// TIA Portal V20 export
// export: Created 2026-10-20T12:50:57.8913211Z, ExportSetting WithDefaults, DisplayName Totally Integrated Automation Portal, DisplayVersion V20 Update 6, DisplayName TIA Portal Openness, DisplayVersion V20 Update 6, DisplayName TIA Portal Version Control Interface, DisplayVersion V20 Update 6, DisplayName SINAMICS Startdrive Advanced, DisplayVersion V20 SP1, DisplayName SINAMICS Startdrive G130, G150, S120, S150, SINAMICS MV, G220, S200, S210, DisplayVersion V20 SP1, DisplayName SINAMICS Startdrive G110M, G120, G120C, G120D, G120P, G115D, DisplayVersion V20 SP1, DisplayName STEP 7 Professional, DisplayVersion V20 Update 6, DisplayName STEP 7 Safety, DisplayVersion V20 Update 2, DisplayName WinCC Basic/Comfort/Advanced, DisplayVersion V20 Update 6, DisplayName WinCC Unified, DisplayVersion V20 Update 6
FUNCTION_BLOCK "Main_Panel"   // FB16, F_LAD
{ S7_Optimized_Access := 'TRUE' }
VERSION : 0.1
// stored: AutoNumber true, IsIECCheckEnabled false, UDAEnableTagReadback false
   VAR_INPUT
      Estop_Cabinet_Ch1 : Bool;
      Reset_Cabinet : Bool;
      Bypass : "F_Bypass_MainPanel";
   END_VAR
   VAR_OUTPUT
      Safety_OK : Bool;
      Main_Panel_OK : Bool;
      Bypass_Warning : Bool;
      ACK { ExternalAccessible := 'False'; ExternalVisible := 'False'; ExternalWritable := 'False'} : Bool;
   END_VAR
   VAR
      Estop_Cabinet_DB : ESTOP1;
   END_VAR
BEGIN

REGION Network 1: RESET CABINET
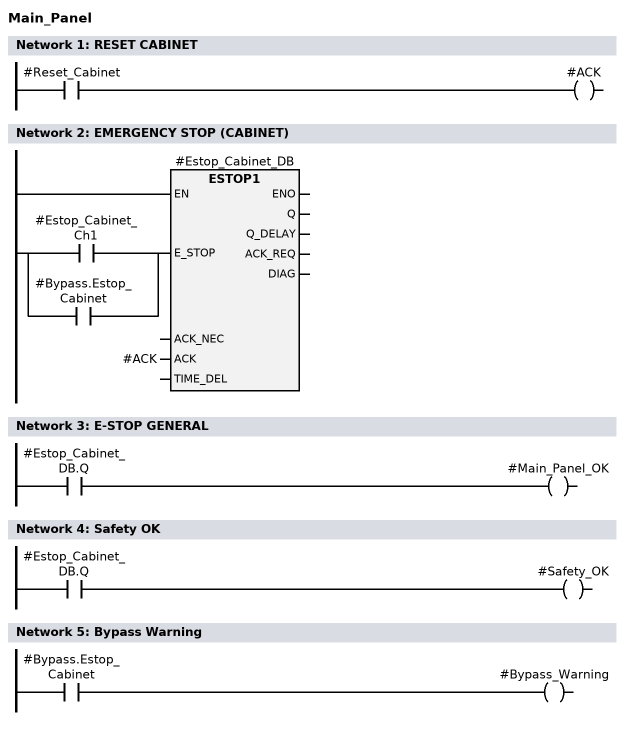
   RUNG wire#powerrail
      Contact( #Reset_Cabinet )
      Coil( #ACK )
   END_RUNG
   // the same network as SCL:
   #ACK := #Reset_Cabinet;
END_REGION

REGION Network 2: EMERGENCY STOP (CABINET)
   RUNG wire#powerrail
      #Estop_Cabinet_DB.ESTOP1(E_STOP := wire#w1, ACK_NEC :=, ACK := #ACK, TIME_DEL :=, Q =>, Q_DELAY =>, ACK_REQ =>, DIAG =>)
   END_RUNG
   RUNG wire#powerrail
      Contact( #Estop_Cabinet_Ch1 )
   END_RUNG wire#w1
   RUNG wire#powerrail
      Contact( #Bypass.Estop_Cabinet )
   END_RUNG wire#w1
   // the same network as SCL:
   #Estop_Cabinet_DB(E_STOP := #Estop_Cabinet_Ch1 OR #Bypass.Estop_Cabinet, ACK := #ACK);   // ESTOP1
END_REGION

REGION Network 3: E-STOP GENERAL
   RUNG wire#powerrail
      Contact( #Estop_Cabinet_DB.Q )
      Coil( #Main_Panel_OK )
   END_RUNG
   // the same network as SCL:
   #Main_Panel_OK := #Estop_Cabinet_DB.Q;
END_REGION

REGION Network 4: Safety OK
   RUNG wire#powerrail
      Contact( #Estop_Cabinet_DB.Q )
      Coil( #Safety_OK )
   END_RUNG
   // the same network as SCL:
   #Safety_OK := #Estop_Cabinet_DB.Q;
END_REGION

REGION Network 5: Bypass Warning
   RUNG wire#powerrail
      Contact( #Bypass.Estop_Cabinet )
      Coil( #Bypass_Warning )
   END_RUNG
   // the same network as SCL:
   #Bypass_Warning := #Bypass.Estop_Cabinet;
END_REGION
END_FUNCTION_BLOCK
